{attribute 'qualified_only'}
{attribute 'strict'}
{attribute 'to_string'}
TYPE E_AxisGeometry : (
    Unknown := 0,
    Linear := 1,
    Rotary := 2
);
END_TYPE

(* stored: Version 1.1.0.1, ProductVersion 3.1.4026.20
   DUT E_AxisGeometry: Id {166dfee1-dc8e-5190-a5fe-022123c3cb66} *)
